{attribute 'qualified_only'}
{attribute 'strict'}
TYPE Platform :
(
	SIMULATION := 0,
	HARDWARE
);
END_TYPE

(* stored: Version 1.1.0.1, ProductVersion 3.1.4026.12
   DUT Platform: Id {fb411fc4-ab63-55e9-b75c-3c8edacd6c24} *)
